FUNCTION_BLOCK PUMP_STATION_LEVEL (* Migrated from IEC 61131-3 ST *)
  (* Standard: 61499-2 *)
  (* Version 1.0, 2026-11-06, st2fb *)
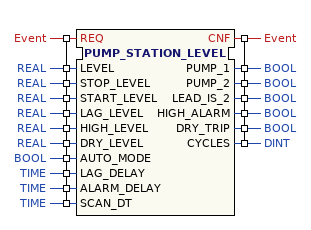
  EVENT_INPUT
    REQ WITH LEVEL, STOP_LEVEL, START_LEVEL, LAG_LEVEL, HIGH_LEVEL, DRY_LEVEL, AUTO_MODE, LAG_DELAY, ALARM_DELAY, SCAN_DT;
  END_EVENT
  EVENT_OUTPUT
    CNF WITH PUMP_1, PUMP_2, LEAD_IS_2, HIGH_ALARM, DRY_TRIP, CYCLES;
  END_EVENT
  VAR_INPUT
    LEVEL : REAL;
    STOP_LEVEL : REAL;
    START_LEVEL : REAL;
    LAG_LEVEL : REAL;
    HIGH_LEVEL : REAL;
    DRY_LEVEL : REAL;
    AUTO_MODE : BOOL;
    LAG_DELAY : TIME;
    ALARM_DELAY : TIME;
    SCAN_DT : TIME;
  END_VAR
  VAR_OUTPUT
    PUMP_1 : BOOL;
    PUMP_2 : BOOL;
    LEAD_IS_2 : BOOL;
    HIGH_ALARM : BOOL;
    DRY_TRIP : BOOL;
    CYCLES : DINT;
  END_VAR
  VAR
    LEAD_REQ : BOOL;
    LAG_REQ : BOOL;
    ST2FB_NOW : TIME;
    LAG_TIMER_IN : BOOL;
    LAG_TIMER_PT : TIME;
    LAG_TIMER_Q : BOOL;
    LAG_TIMER_ET : TIME;
    LAG_TIMER_STATE : INT;
    LAG_TIMER_PREV_IN : BOOL;
    LAG_TIMER_START_TIME : TIME;
    ALARM_TIMER_IN : BOOL;
    ALARM_TIMER_PT : TIME;
    ALARM_TIMER_Q : BOOL;
    ALARM_TIMER_ET : TIME;
    ALARM_TIMER_STATE : INT;
    ALARM_TIMER_PREV_IN : BOOL;
    ALARM_TIMER_START_TIME : TIME;
    LEAD_STOPPED_CLK : BOOL;
    LEAD_STOPPED_Q : BOOL;
    LEAD_STOPPED_M : BOOL;
  END_VAR
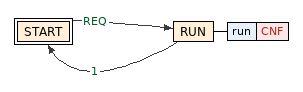
  EC_STATES
    START;
    RUN : run -> CNF;
  END_STATES
  EC_TRANSITIONS
    START TO RUN := REQ;
    RUN TO START := 1;
  END_TRANSITIONS
  ALGORITHM run IN ST:
ST2FB_NOW := ST2FB_NOW + SCAN_DT;
DRY_TRIP := LEVEL <= DRY_LEVEL;
IF NOT AUTO_MODE OR DRY_TRIP OR LEVEL <= STOP_LEVEL THEN
  LEAD_REQ := FALSE;
ELSIF LEVEL >= START_LEVEL THEN
  LEAD_REQ := TRUE;
END_IF;

LAG_TIMER_IN := LEAD_REQ AND LEVEL >= LAG_LEVEL;
LAG_TIMER_PT := LAG_DELAY;
IF (LAG_TIMER_STATE = 0) AND NOT LAG_TIMER_PREV_IN AND LAG_TIMER_IN THEN
  LAG_TIMER_STATE := 1;
  LAG_TIMER_Q := FALSE;
  LAG_TIMER_START_TIME := ST2FB_NOW;
ELSE
  IF NOT LAG_TIMER_IN THEN
    LAG_TIMER_ET := T#0s;
    LAG_TIMER_Q := FALSE;
    LAG_TIMER_STATE := 0;
  ELSIF LAG_TIMER_STATE = 1 THEN
    IF LAG_TIMER_START_TIME + LAG_TIMER_PT <= ST2FB_NOW THEN
      LAG_TIMER_STATE := 2;
      LAG_TIMER_Q := TRUE;
      LAG_TIMER_ET := LAG_TIMER_PT;
    ELSE
      LAG_TIMER_ET := ST2FB_NOW - LAG_TIMER_START_TIME;
    END_IF;
  END_IF;
END_IF;
LAG_TIMER_PREV_IN := LAG_TIMER_IN;

IF NOT LEAD_REQ THEN
  LAG_REQ := FALSE;
ELSIF LAG_TIMER_Q THEN
  LAG_REQ := TRUE;
END_IF;

LEAD_STOPPED_CLK := LEAD_REQ;
LEAD_STOPPED_Q := NOT LEAD_STOPPED_CLK AND NOT LEAD_STOPPED_M;
LEAD_STOPPED_M := NOT LEAD_STOPPED_CLK;

IF LEAD_STOPPED_Q THEN
  LEAD_IS_2 := NOT LEAD_IS_2;
  CYCLES := CYCLES + 1;
END_IF;
IF LEAD_IS_2 THEN
  PUMP_2 := LEAD_REQ;
  PUMP_1 := LAG_REQ;
ELSE
  PUMP_1 := LEAD_REQ;
  PUMP_2 := LAG_REQ;
END_IF;

ALARM_TIMER_IN := LEVEL >= HIGH_LEVEL;
ALARM_TIMER_PT := ALARM_DELAY;
IF (ALARM_TIMER_STATE = 0) AND NOT ALARM_TIMER_PREV_IN AND ALARM_TIMER_IN THEN
  ALARM_TIMER_STATE := 1;
  ALARM_TIMER_Q := FALSE;
  ALARM_TIMER_START_TIME := ST2FB_NOW;
ELSE
  IF NOT ALARM_TIMER_IN THEN
    ALARM_TIMER_ET := T#0s;
    ALARM_TIMER_Q := FALSE;
    ALARM_TIMER_STATE := 0;
  ELSIF ALARM_TIMER_STATE = 1 THEN
    IF ALARM_TIMER_START_TIME + ALARM_TIMER_PT <= ST2FB_NOW THEN
      ALARM_TIMER_STATE := 2;
      ALARM_TIMER_Q := TRUE;
      ALARM_TIMER_ET := ALARM_TIMER_PT;
    ELSE
      ALARM_TIMER_ET := ST2FB_NOW - ALARM_TIMER_START_TIME;
    END_IF;
  END_IF;
END_IF;
ALARM_TIMER_PREV_IN := ALARM_TIMER_IN;
HIGH_ALARM := ALARM_TIMER_Q;
  END_ALGORITHM
END_FUNCTION_BLOCK
